Fanuc KAREL source: KX00027.KL

PROGRAM KX00027
%NOLOCKGROUP
%STACKSIZE = 1000
VAR
  I: INTEGER
  J: INTEGER
  B: BOOLEAN
  F: FILE
  S: STRING[80]
  P: XYZWPR
BEGIN
  I = 1
END KX00027
